Yaskawa INFORM job: 1-DEFRO-5-KOSZ.JBI

/JOB
//NAME 1-DEFRO-5-KOSZ
//POS
///NPOS 37,37,37,0,0,0
///TOOL 0
///POSTYPE PULSE
///PULSE
C00000=-283,-101162,-84213,3710,-80188,-1936
C00001=-275,-97864,-82985,3720,-79251,-1967
C00002=-100003,31603,4033,-7680,-72698,-47529
C00003=-100001,31607,4031,-7680,-72698,-47532
C00004=-101284,101717,15156,-4078,-52370,-88533
C00005=-106030,98783,11088,-3548,-51538,-87057
C00006=-101741,79318,-156,-3344,-46518,35055
C00007=-103126,90079,-944,-3752,-40557,35773
C00008=-103126,90079,-944,-3752,-40557,35773
C00009=-103831,97844,9734,-3579,-43155,35906
C00010=-102596,65773,-9481,200,-39522,35767
C00011=-102596,65773,-9481,6832,-44909,-46607
C00012=-97155,78202,-19745,30250,-25050,-62284
C00013=-98162,85024,-10279,27721,-26879,-60727
C00014=-96622,56300,-24733,23618,-32509,-59065
C00015=-96079,53622,-29140,32876,-19135,-23317
C00016=-95299,74134,-28399,77084,-12548,-43279
C00017=-101099,71014,-32620,83437,-10098,-44474
C00018=-101099,52121,-34889,47023,-13961,-27940
C00019=-101099,36619,-33203,29323,-21209,-19692
C00020=-101099,36619,-33203,29323,-21209,-19692
C00021=-101801,67266,-42312,144719,-12916,-72337
C00022=-95588,69918,-38485,130896,-13770,-67922
C00023=-95035,59333,-32585,57682,-14738,-34474
C00024=-94481,79102,-16755,23606,-29701,-18576
C00025=-99899,75728,-21276,23527,-27793,-16866
C00026=-99086,45522,-41235,42765,-18284,-25961
C00027=-100543,55433,-28857,2241,-34808,32636
C00028=-107763,109938,23476,-14806,-64763,39357
C00029=-107254,101652,11557,-15338,-61720,39618
C00030=-107352,87208,9990,-14558,-67984,38821
C00031=-98885,97187,8635,10637,-50243,-42045
C00032=-97889,89767,-1552,10913,-47920,-42616
C00033=-97858,62636,-1557,9208,-61662,-41293
C00034=-100003,31603,4033,-7680,-72698,-47529
C00035=-275,-97864,-82985,3720,-79251,-1967
C00036=-283,-101162,-84213,3710,-80188,-1936
BC00000=570125
BC00001=808681
BC00002=808681
BC00003=808680
BC00004=808680
BC00005=808680
BC00006=808680
BC00007=808680
BC00008=808680
BC00009=808680
BC00010=808680
BC00011=808680
BC00012=808680
BC00013=808680
BC00014=808680
BC00015=808680
BC00016=808680
BC00017=808680
BC00018=808680
BC00019=808680
BC00020=808680
BC00021=808680
BC00022=808680
BC00023=808679
BC00024=808679
BC00025=808679
BC00026=808679
BC00027=808679
BC00028=808679
BC00029=808679
BC00030=808679
BC00031=808679
BC00032=808679
BC00033=808679
BC00034=808681
BC00035=808681
BC00036=570125
EC00000=1,-94526
EC00001=1,-94526
EC00002=1,-94526
EC00003=119163,-211743
EC00004=119163,-212879
EC00005=119163,-212879
EC00006=119163,-212879
EC00007=119163,-212879
EC00008=119163,-212879
EC00009=119163,-212879
EC00010=119163,-211743
EC00011=119163,-211743
EC00012=119163,-211743
EC00013=119163,-211743
EC00014=119163,-211743
EC00015=119163,-211743
EC00016=119163,-211743
EC00017=119163,-211743
EC00018=119163,-211743
EC00019=119163,167367
EC00020=119163,167367
EC00021=119163,167367
EC00022=119164,167366
EC00023=119163,167367
EC00024=119163,167367
EC00025=119163,167367
EC00026=119163,167367
EC00027=119163,167367
EC00028=119163,167367
EC00029=119163,167367
EC00030=119163,167367
EC00031=119163,167367
EC00032=119163,167367
EC00033=119163,167367
EC00034=1,-94526
EC00035=1,-94526
EC00036=1,-94526
//INST
///DATE 2025/01/14 11:01
///ATTR SC,RW
///GROUP1 RB1,BS1
///GROUP2 ST3
NOP
MOVJ C00000 BC00000 VJ=40.00 DEC=20  +MOVJ EC00000 VJ=40.00
MOVJ C00001 BC00001 VJ=40.00 DEC=20  +MOVJ EC00001 VJ=40.00
MOVJ C00002 BC00002 VJ=40.00 DEC=20  +MOVJ EC00002 VJ=40.00
MOVJ C00003 BC00003 VJ=20.00 DEC=20  +MOVJ EC00003 VJ=20.00
MOVJ C00004 BC00004 VJ=20.00 DEC=20  +MOVJ EC00004 VJ=20.00
MACRO1 MJ#(0) ARGF5
ARCON
MOVL C00005 BC00005 V=4.2 DEC=20  +MOVJ EC00005 VJ=20.00
ARCOF
MOVJ C00006 BC00006 VJ=20.00 DEC=20  +MOVJ EC00006 VJ=20.00
MOVJ C00007 BC00007 VJ=20.00 DEC=20  +MOVJ EC00007 VJ=20.00
MOVJ C00008 BC00008 VJ=20.00 DEC=20  +MOVJ EC00008 VJ=20.00
ARCON
MOVL C00009 BC00009 V=4.2 DEC=20  +MOVJ EC00009 VJ=20.00
ARCOF
MOVJ C00010 BC00010 VJ=20.00 DEC=20  +MOVJ EC00010 VJ=20.00
MOVJ C00011 BC00011 VJ=20.00 DEC=20  +MOVJ EC00011 VJ=20.00
MOVJ C00012 BC00012 VJ=20.00 DEC=20  +MOVJ EC00012 VJ=20.00
ARCON
MOVL C00013 BC00013 V=4.2 DEC=20  +MOVJ EC00013 VJ=20.00
ARCOF
MOVJ C00014 BC00014 VJ=20.00 DEC=20  +MOVJ EC00014 VJ=20.00
MOVJ C00015 BC00015 VJ=20.00 DEC=20  +MOVJ EC00015 VJ=20.00
MOVJ C00016 BC00016 VJ=30.00 DEC=20  +MOVJ EC00016 VJ=0.78
ARCON
WVON WEV#(1)
MOVL C00017 BC00017 V=4.2 DEC=20  +MOVJ EC00017 VJ=0.78
WVOF
ARCOF
MOVJ C00018 BC00018 VJ=30.00 DEC=20  +MOVJ EC00018 VJ=30.00
MOVJ C00019 BC00019 VJ=40.00 DEC=20  +MOVJ EC00019 VJ=30.00
MOVJ C00020 BC00020 VJ=40.00 DEC=20  +MOVJ EC00020 VJ=30.00
MOVJ C00021 BC00021 VJ=30.00 DEC=20  +MOVJ EC00021 VJ=30.00
ARCON
WVON WEV#(1)
MOVL C00022 BC00022 V=4.2 DEC=20  +MOVJ EC00022 VJ=30.00
WVOF
ARCOF
MOVJ C00023 BC00023 VJ=30.00 DEC=20  +MOVJ EC00023 VJ=30.00
MOVJ C00024 BC00024 VJ=30.00 DEC=20  +MOVJ EC00024 VJ=30.00
ARCON
MOVL C00025 BC00025 V=4.2 DEC=20  +MOVJ EC00025 VJ=30.00
ARCOF
MOVJ C00026 BC00026 VJ=30.00 DEC=20  +MOVJ EC00026 VJ=30.00
MOVJ C00027 BC00027 VJ=30.00 DEC=20  +MOVJ EC00027 VJ=30.00
MOVJ C00028 BC00028 VJ=30.00 DEC=20  +MOVJ EC00028 VJ=30.00
ARCON
MOVL C00029 BC00029 V=4.2 DEC=20  +MOVJ EC00029 VJ=30.00
ARCOF
MOVJ C00030 BC00030 VJ=30.00 DEC=20  +MOVJ EC00030 VJ=30.00
MOVJ C00031 BC00031 VJ=30.00 DEC=20  +MOVJ EC00031 VJ=30.00
ARCON
MOVL C00032 BC00032 V=4.2 DEC=20  +MOVJ EC00032 VJ=30.00
ARCOF
MOVJ C00033 BC00033 VJ=30.00 DEC=20  +MOVJ EC00033 VJ=30.00
MOVJ C00034 BC00034 VJ=30.00 DEC=20  +MOVJ EC00034 VJ=30.00
MOVJ C00035 BC00035 VJ=30.00 DEC=20  +MOVJ EC00035 VJ=30.00
MOVJ C00036 BC00036 VJ=30.00 DEC=20  +MOVJ EC00036 VJ=30.00
END
